FUNCTION_BLOCK IO_GUARD (* Migrated from IEC 61131-3 ST *)
  (* Standard: 61499-2 *)
  (* Version 1.0, 2026-11-06, st2fb *)
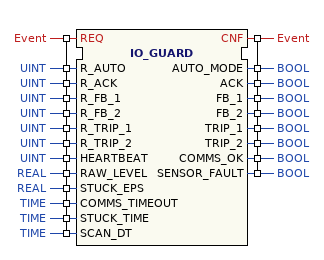
  EVENT_INPUT
    REQ WITH R_AUTO, R_ACK, R_FB_1, R_FB_2, R_TRIP_1, R_TRIP_2, HEARTBEAT, RAW_LEVEL, STUCK_EPS, COMMS_TIMEOUT, STUCK_TIME, SCAN_DT;
  END_EVENT
  EVENT_OUTPUT
    CNF WITH AUTO_MODE, ACK, FB_1, FB_2, TRIP_1, TRIP_2, COMMS_OK, SENSOR_FAULT;
  END_EVENT
  VAR_INPUT
    R_AUTO : UINT;
    R_ACK : UINT;
    R_FB_1 : UINT;
    R_FB_2 : UINT;
    R_TRIP_1 : UINT;
    R_TRIP_2 : UINT;
    HEARTBEAT : UINT;
    RAW_LEVEL : REAL;
    STUCK_EPS : REAL;
    COMMS_TIMEOUT : TIME;
    STUCK_TIME : TIME;
    SCAN_DT : TIME;
  END_VAR
  VAR_OUTPUT
    AUTO_MODE : BOOL;
    ACK : BOOL;
    FB_1 : BOOL;
    FB_2 : BOOL;
    TRIP_1 : BOOL;
    TRIP_2 : BOOL;
    COMMS_OK : BOOL;
    SENSOR_FAULT : BOOL;
  END_VAR
  VAR
    LAST_HEARTBEAT : UINT;
    LAST_LEVEL : REAL;
    SEEN_BEAT : BOOL;
    UNCHANGED : BOOL;
    DELTA : REAL;
    ST2FB_NOW : TIME;
    COMMS_TIMER_IN : BOOL;
    COMMS_TIMER_PT : TIME;
    COMMS_TIMER_Q : BOOL;
    COMMS_TIMER_ET : TIME;
    COMMS_TIMER_STATE : INT;
    COMMS_TIMER_PREV_IN : BOOL;
    COMMS_TIMER_START_TIME : TIME;
    STUCK_TIMER_IN : BOOL;
    STUCK_TIMER_PT : TIME;
    STUCK_TIMER_Q : BOOL;
    STUCK_TIMER_ET : TIME;
    STUCK_TIMER_STATE : INT;
    STUCK_TIMER_PREV_IN : BOOL;
    STUCK_TIMER_START_TIME : TIME;
    ACK_EDGE_CLK : BOOL;
    ACK_EDGE_Q : BOOL;
    ACK_EDGE_M : BOOL;
    FAULT_LATCH_S1 : BOOL;
    FAULT_LATCH_R : BOOL;
    FAULT_LATCH_Q1 : BOOL;
  END_VAR
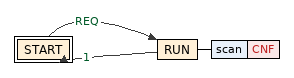
  EC_STATES
    START;
    RUN : scan -> CNF;
  END_STATES
  EC_TRANSITIONS
    START TO RUN := REQ;
    RUN TO START := 1;
  END_TRANSITIONS
  ALGORITHM scan IN ST:
ST2FB_NOW := ST2FB_NOW + SCAN_DT;
IF HEARTBEAT <> LAST_HEARTBEAT THEN
  SEEN_BEAT := TRUE;
END_IF;
COMMS_TIMER_IN := HEARTBEAT = LAST_HEARTBEAT;
COMMS_TIMER_PT := COMMS_TIMEOUT;
IF COMMS_TIMER_STATE = 0 AND NOT COMMS_TIMER_PREV_IN AND COMMS_TIMER_IN THEN
  COMMS_TIMER_STATE := 1;
  COMMS_TIMER_Q := FALSE;
  COMMS_TIMER_START_TIME := ST2FB_NOW;
ELSE
  IF NOT COMMS_TIMER_IN THEN
    COMMS_TIMER_ET := T#0s;
    COMMS_TIMER_Q := FALSE;
    COMMS_TIMER_STATE := 0;
  ELSIF COMMS_TIMER_STATE = 1 THEN
    IF COMMS_TIMER_START_TIME + COMMS_TIMER_PT <= ST2FB_NOW THEN
      COMMS_TIMER_STATE := 2;
      COMMS_TIMER_Q := TRUE;
      COMMS_TIMER_ET := COMMS_TIMER_PT;
    ELSE
      COMMS_TIMER_ET := ST2FB_NOW - COMMS_TIMER_START_TIME;
    END_IF;
  END_IF;
END_IF;
COMMS_TIMER_PREV_IN := COMMS_TIMER_IN;
LAST_HEARTBEAT := HEARTBEAT;
COMMS_OK := SEEN_BEAT AND NOT COMMS_TIMER_Q;
DELTA := RAW_LEVEL - LAST_LEVEL;
UNCHANGED := DELTA <= STUCK_EPS AND DELTA >= -STUCK_EPS;
LAST_LEVEL := RAW_LEVEL;
STUCK_TIMER_IN := UNCHANGED AND COMMS_OK;
STUCK_TIMER_PT := STUCK_TIME;
IF STUCK_TIMER_STATE = 0 AND NOT STUCK_TIMER_PREV_IN AND STUCK_TIMER_IN THEN
  STUCK_TIMER_STATE := 1;
  STUCK_TIMER_Q := FALSE;
  STUCK_TIMER_START_TIME := ST2FB_NOW;
ELSE
  IF NOT STUCK_TIMER_IN THEN
    STUCK_TIMER_ET := T#0s;
    STUCK_TIMER_Q := FALSE;
    STUCK_TIMER_STATE := 0;
  ELSIF STUCK_TIMER_STATE = 1 THEN
    IF STUCK_TIMER_START_TIME + STUCK_TIMER_PT <= ST2FB_NOW THEN
      STUCK_TIMER_STATE := 2;
      STUCK_TIMER_Q := TRUE;
      STUCK_TIMER_ET := STUCK_TIMER_PT;
    ELSE
      STUCK_TIMER_ET := ST2FB_NOW - STUCK_TIMER_START_TIME;
    END_IF;
  END_IF;
END_IF;
STUCK_TIMER_PREV_IN := STUCK_TIMER_IN;
ACK := R_ACK <> 0;
ACK_EDGE_CLK := ACK;
ACK_EDGE_Q := ACK_EDGE_CLK AND NOT ACK_EDGE_M;
ACK_EDGE_M := ACK_EDGE_CLK;
FAULT_LATCH_S1 := STUCK_TIMER_Q;
FAULT_LATCH_R := ACK_EDGE_Q;
FAULT_LATCH_Q1 := FAULT_LATCH_S1 OR NOT FAULT_LATCH_R AND FAULT_LATCH_Q1;
SENSOR_FAULT := FAULT_LATCH_Q1;
AUTO_MODE := R_AUTO <> 0 AND COMMS_OK AND NOT SENSOR_FAULT;
FB_1 := R_FB_1 <> 0;
FB_2 := R_FB_2 <> 0;
TRIP_1 := R_TRIP_1 <> 0;
TRIP_2 := R_TRIP_2 <> 0;
  END_ALGORITHM
END_FUNCTION_BLOCK
